FUNCTION_BLOCK Sorting (* Composite Function Block Type *)
  (* Standard: 61499-2 *)
  (* Version 0.0, 7/2/2026, template *)
  PACKAGE Main;
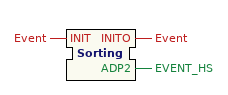
  EVENT_INPUT
    INIT; (* Initialization Request *)
  END_EVENT
  EVENT_OUTPUT
    INITO; (* Initialization Confirm *)
  END_EVENT
  PLUGS
    ADP2 : EVENT_HS;
  END_PLUGS
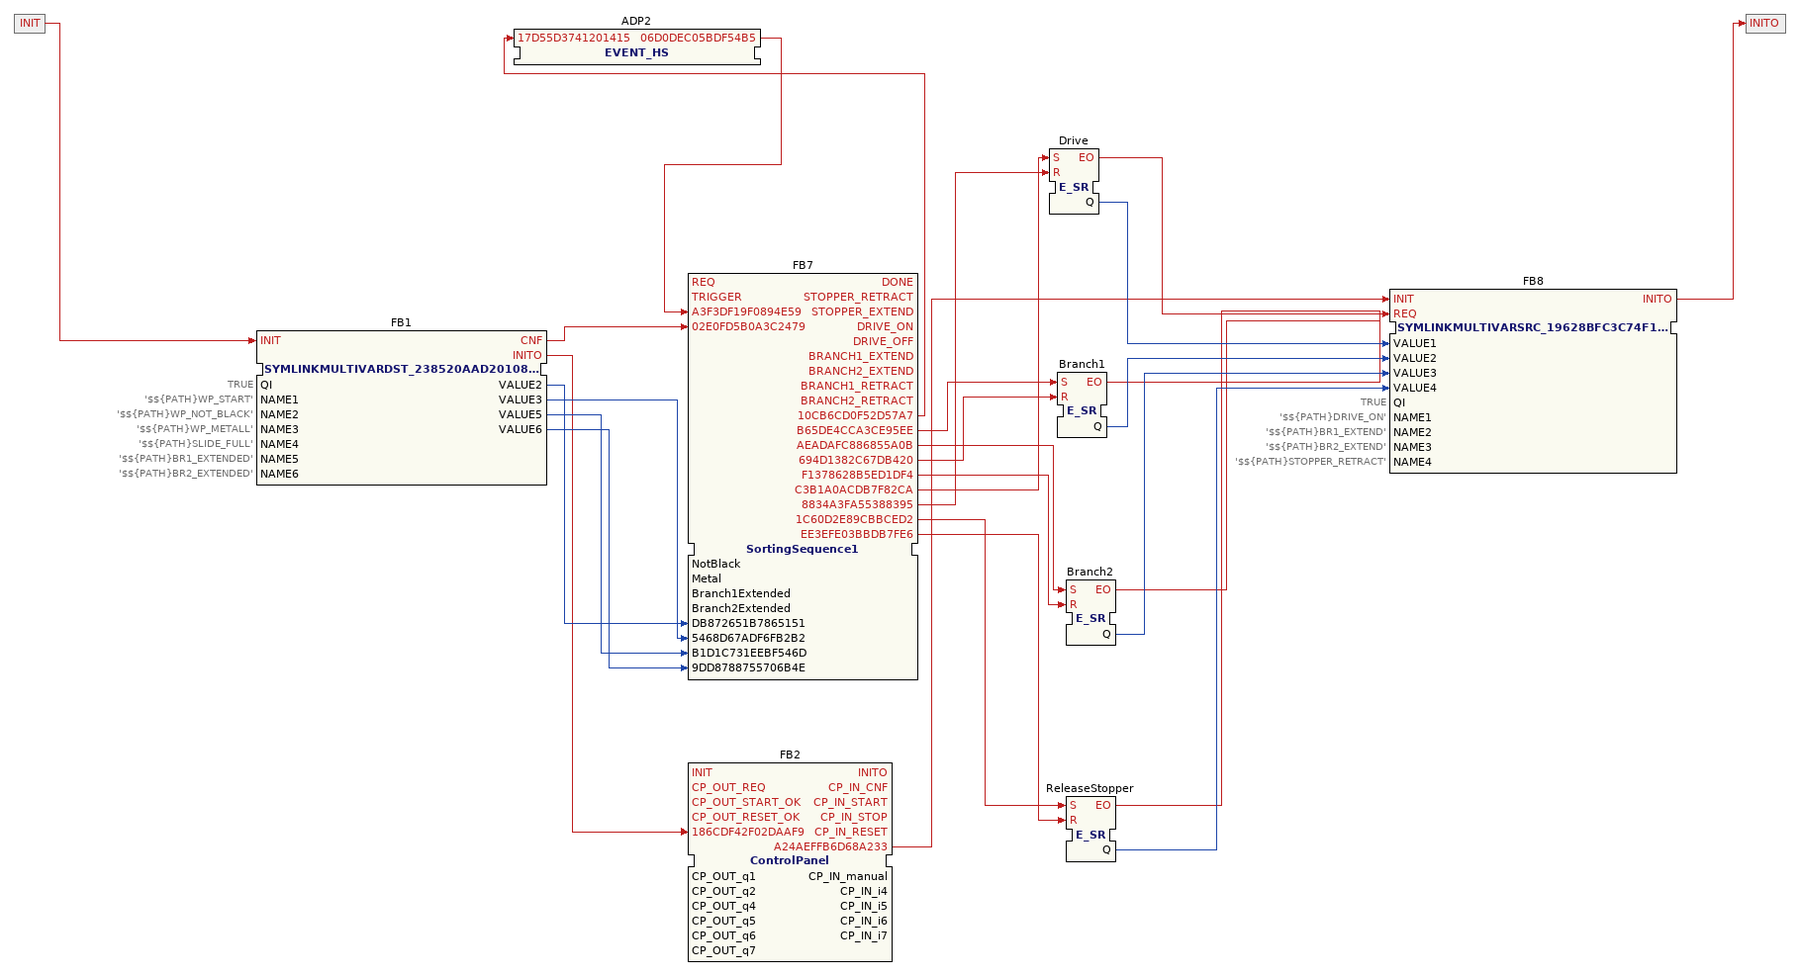
  FBS
    FB1 : SYMLINKMULTIVARDST_238520AAD20108C65(QI := TRUE, NAME1 := '$${PATH}WP_START', NAME2 := '$${PATH}WP_NOT_BLACK', NAME3 := '$${PATH}WP_METALL', NAME4 := '$${PATH}SLIDE_FULL', NAME5 := '$${PATH}BR1_EXTENDED', NAME6 := '$${PATH}BR2_EXTENDED'); {SET_ATTRIBUTE(Configuration.GenericFBType.InterfaceParams, Runtime.System#I:=7;VALUE${I$}:BOOL,BOOL,BOOL,BOOL,BOOL,BOOL,BOOL)}
    FB2 : ControlPanel;
    Drive : E_SR;
    Branch1 : E_SR;
    Branch2 : E_SR;
    ReleaseStopper : E_SR;
    FB7 : SortingSequence1;
    FB8 : SYMLINKMULTIVARSRC_19628BFC3C74F1AB1(QI := TRUE, NAME1 := '$${PATH}DRIVE_ON', NAME2 := '$${PATH}BR1_EXTEND', NAME3 := '$${PATH}BR2_EXTEND', NAME4 := '$${PATH}STOPPER_RETRACT'); {SET_ATTRIBUTE(Configuration.GenericFBType.InterfaceParams, Runtime.System#I:=4;VALUE${I$}:BOOL,BOOL,BOOL,BOOL)}
  END_FBS
  EVENT_CONNECTIONS
    INIT TO FB1.INIT;
    ADP2.06D0DEC05BDF54B5 TO FB7.A3F3DF19F0894E59;
    FB1.CNF TO FB7.02E0FD5B0A3C2479;
    FB1.INITO TO FB2.186CDF42F02DAAF9;
    FB7.10CB6CD0F52D57A7 TO ADP2.17D55D3741201415;
    FB2.A24AEFFB6D68A233 TO FB8.INIT;
    FB8.INITO TO INITO;
    Drive.EO TO FB8.REQ;
    Branch1.EO TO FB8.REQ;
    Branch2.EO TO FB8.REQ;
    ReleaseStopper.EO TO FB8.REQ;
    FB7.B65DE4CCA3CE95EE TO Branch1.S;
    FB7.AEADAFC886855A0B TO Branch2.S;
    FB7.694D1382C67DB420 TO Branch1.R;
    FB7.F1378628B5ED1DF4 TO Branch2.R;
    FB7.C3B1A0ACDB7F82CA TO Drive.S;
    FB7.8834A3FA55388395 TO Drive.R;
    FB7.1C60D2E89CBBCED2 TO ReleaseStopper.S;
    FB7.EE3EFE03BBDB7FE6 TO ReleaseStopper.R;
  END_CONNECTIONS
  DATA_CONNECTIONS
    FB1.VALUE2 TO FB7.DB872651B7865151;
    FB1.VALUE3 TO FB7.5468D67ADF6FB2B2;
    FB1.VALUE5 TO FB7.B1D1C731EEBF546D;
    FB1.VALUE6 TO FB7.9DD8788755706B4E;
    Drive.Q TO FB8.VALUE1;
    Branch1.Q TO FB8.VALUE2;
    Branch2.Q TO FB8.VALUE3;
    ReleaseStopper.Q TO FB8.VALUE4;
  END_CONNECTIONS
END_FUNCTION_BLOCK
